FUNCTION_BLOCK TankValves (* Basic Function Block Type *)
  (* Standard: 61499-2 *)
  (* Version 0.0, 6/20/2016, Andrei, nxtControl GmbH, Template *)
  PACKAGE Main;
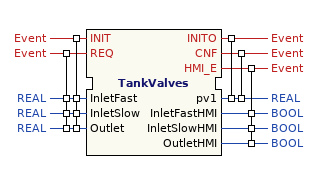
  EVENT_INPUT
    INIT WITH InletFast, InletSlow, Outlet; (* Initialization Request *)
    REQ WITH InletFast, InletSlow, Outlet; (* Normal Execution Request *)
  END_EVENT
  EVENT_OUTPUT
    INITO WITH pv1; (* Initialization Confirm *)
    CNF WITH pv1; (* Execution Confirmation *)
    HMI_E WITH InletFastHMI, InletSlowHMI, OutletHMI;
  END_EVENT
  VAR_INPUT
    InletFast : REAL; (* Input event qualifier *)
    InletSlow : REAL;
    Outlet : REAL;
  END_VAR
  VAR_OUTPUT
    pv1 : REAL; (* Output event qualifier *)
    InletFastHMI : BOOL;
    InletSlowHMI : BOOL;
    OutletHMI : BOOL;
  END_VAR
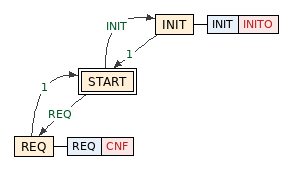
  EC_STATES
    START; (* Initial State *)
    INIT : INIT -> INITO; (* Initialization *)
    REQ : REQ -> CNF; (* Normal execution *)
  END_STATES
  EC_TRANSITIONS
    START TO INIT := INIT;
    INIT TO START := 1;
    START TO REQ := REQ;
    REQ TO START := 1;
  END_TRANSITIONS
  ALGORITHM INIT IN ST: (* Initialization algorithm *)
pv1 := 0.0;;
  END_ALGORITHM
  ALGORITHM REQ IN ST: (* Normally executed algorithm *)
pv1 := 200.0*(InletFast) + 100.0*(InletSlow) -150.0 * (Outlet);


InletFastHMI := INT_TO_BOOL(REAL_TO_INT(InletFast));
InletSlowHMI := INT_TO_BOOL(REAL_TO_INT(InletSlow));
OutletHMI := INT_TO_BOOL(REAL_TO_INT(Outlet));
  END_ALGORITHM
END_FUNCTION_BLOCK
